// This function has been automatically generated from the project information.
{attribute 'signature_flag' := '1073741824'}
{attribute 'TcGenerated'}
{attribute 'no-analysis'}
FUNCTION F_GetTitle : WSTRING
VAR_INPUT
	
END_VAR

F_GetTitle := "PersistentDataHandler";

END_FUNCTION

(* stored: Version 1.1.0.1
   POU F_GetTitle: Id {8ab97be1-a88f-486f-a7fc-9852ca980e0b}, SpecialFunc None *)
